Fanuc KAREL source: ke00002.KL

-- PROVISIONAL review KL for V770-1; original PC SHA256 da65d6fe0206fb9efbb06fc4987a072e8940dec7b978e8dd12ac78c5eefaa3cf
-- Incomplete behavior may be omitted. Consult companion uncertainty JSON. Do not deploy.
PROGRAM KE00002
%NOLOCKGROUP
BEGIN
  -- UNRESOLVED_PC offsets 5-17; opcodes 3F,75
  -- UNRESOLVED_PC offsets 22-29; opcodes 9D,23
  -- UNRESOLVED_PC offsets 34-46; opcodes 3F,22,9D,33,61
  -- UNRESOLVED_PC offsets 51-87; opcodes 27,22,2A,22,22,22,22,31
  -- UNRESOLVED_PC offsets 92-96; opcodes 7F
END KE00002
